(*
	A pump skid's status, read by the master from the skid's GVL.status over ADS. A command has
	settled when sequence matches the command's and busy is clear.
	Keep this identical to ST_SkidStatus in every skid project: ADS copies it byte for byte.
*)
TYPE ST_SkidStatus :
STRUCT
	sequence: UDINT;  // the last command the skid accepted
	busy: BOOL;  // staging up or down, until the skid's staging span has ended
	running: BOOL;  // staged up
	faulted: BOOL;  // the last command ended in a fault
	faultText: STRING(80);  // why, when faulted
	flowRate: REAL;  // GPM
END_STRUCT
END_TYPE

(* stored: Version 1.1.0.1
   DUT ST_SkidStatus: Id {c0e86fad-b726-4363-b806-bd6fb12e327b} *)
